FUNCTION_BLOCK FB_Valve
VAR_INPUT
    bOpen : BOOL;
END_VAR
VAR_OUTPUT
    bIsOpen : BOOL;
END_VAR

bIsOpen := bOpen;
	bIsOpen := NOT bOpen;
bOpen := FALSE;

END_FUNCTION_BLOCK

(* stored: Version 1.1.0.1, ProductVersion 3.1.4024.12
   POU FB_Valve: Id {11111111-2222-3333-4444-555555555557}, SpecialFunc None *)
